Staubli VAL3: robotStatus.pgx

public program robotStatus()
begin
  //检测状态显示变化
  if _sRobotStatus!=sLstRobStatus
    sLstRobStatus=_sRobotStatus
    call Log:addlog(toString(".3",clock())+" "+"[状态信息]:"+_sRobotStatus+getDate(" %m-%d %H:%M:%S"),1)
  endIf

  if sTrajStatus!=sLstTrajStatus
    sLstTrajStatus=sTrajStatus
    call Log:addlog(toString(".3",clock())+" "+"[路径信息]:"+sTrajStatus+getDate(" %m-%d %H:%M:%S"),2)
  endIf

  if sIOStatus!=sLstIOStatus
    sLstIOStatus=sIOStatus
    call Log:addlog(toString(".3",clock())+" "+"[信号信息]:"+sIOStatus+getDate(" %m-%d %H:%M:%S"),3)
  endIf
end
